(* IEC 61131-3 sources: tsplc/examples/bottling-line/raw-st/src/io, 2 files *)

(* ---- IO.st ---- *)
{attribute 'qualified_only'}
VAR_GLOBAL
	StartButton : BOOL;
	BottlePresent : BOOL;
	CapperRun : BOOL;
	ZoneStatus : UINT;
	InfeedSpeed : UINT;
END_VAR

(* ---- PRG_ReadInputs.st ---- *)
PROGRAM PRG_ReadInputs
VAR
	Cycles : UDINT;
END_VAR
Cycles := Cycles + 1;
END_PROGRAM
